FUNCTION_BLOCK FB_PendantErrorState EXTENDS FB_PendantState
VAR_INPUT
END_VAR
VAR_OUTPUT
END_VAR
VAR
END_VAR

METHOD ResetCommand : BOOL
pPendant^._Error := FALSE;
pPendant^.SetState(pPendant^.fbPendantPreInitState);
END_METHOD


METHOD RunState : BOOL
ResetCommand();
END_METHOD

PROPERTY StateID : STRING
GET
StateID := 'Error State';
END_GET
END_PROPERTY

END_FUNCTION_BLOCK

(* stored: Version 1.1.0.1, ProductVersion 3.1.4024.15
   POU FB_PendantErrorState: Id {b58925e1-a00e-4433-a211-7c74b6d09ad0}, SpecialFunc None
   Method ResetCommand: Id {d4a76690-9e3b-4a78-8d7d-85736c716d0c}
   Method RunState: Id {90673749-d9e7-445a-b04c-e1d5d49f143d}
   Property StateID: Id {85f67b1d-627d-4ee1-8811-980e6bac68d4}
   Get Get: Id {c08cbac7-562a-4d90-89bf-3396f2fdc2f4} *)
